Staubli VAL3: pointEdit.pgx

public program pointEdit()
  local bool l_bExit
begin

end
